// TIA Portal V20 export
Screen "Pop-up_VISION OFFSET VALUES"  395x635
  ScreenItem "Robot Name" at 2,2 size 393x48  Type=HmiIOField
  ScreenItem "Background" at -1,49 size 395x586  Type=HmiRectangle
  ScreenItem "Cancel Mode" at 315,4 size 76x42  Type=HmiButton
  ScreenItem "矩形_4" at 9,62 size 378x540  Type=HmiRectangle
  ScreenItem "Text field Robot Status_5" at 9,63 size 378x30  Type=HmiTextBox
  ScreenItem "FaultNo" at 251,99 size 108x63  Type=HmiIOField
  ScreenItem "Text field_8" at 20,117 size 223x29  Type=HmiTextBox
  ScreenItem "Text field_1" at 20,195 size 223x29  Type=HmiTextBox
  ScreenItem "FaultNo_1" at 251,176 size 108x63  Type=HmiIOField
  ScreenItem "FaultNo_2" at 250,331 size 108x63  Type=HmiIOField
  ScreenItem "Text field_2" at 19,350 size 223x29  Type=HmiTextBox
  ScreenItem "Text field_3" at 19,272 size 223x29  Type=HmiTextBox
  ScreenItem "FaultNo_3" at 250,254 size 108x63  Type=HmiIOField
  ScreenItem "FaultNo_4" at 250,495 size 108x63  Type=HmiIOField
  ScreenItem "Text field_4" at 19,514 size 223x29  Type=HmiTextBox
  ScreenItem "Text field_5" at 19,436 size 223x29  Type=HmiTextBox
  ScreenItem "FaultNo_5" at 250,418 size 108x63  Type=HmiIOField
